FUNCTION_BLOCK Agua_Reuso_HMI (* Service Interface Function Block Type *)
  (* Standard: 61499-2 *)
  (* Version 1.2, 15/10/2026, Hidryco, Hidryco, IHM da Agua_Reuso *)
  PACKAGE Hidryco.HidrycoLib;
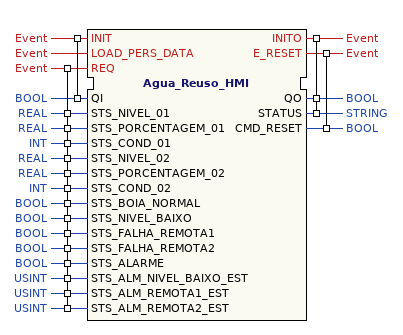
  EVENT_INPUT
    INIT WITH QI;
    LOAD_PERS_DATA; (* Reenvia os parametros persistentes *)
    REQ WITH STS_NIVEL_01, STS_PORCENTAGEM_01, STS_COND_01, STS_NIVEL_02, STS_PORCENTAGEM_02, STS_COND_02, STS_BOIA_NORMAL, STS_NIVEL_BAIXO, STS_FALHA_REMOTA1, STS_FALHA_REMOTA2, STS_ALARME, STS_ALM_NIVEL_BAIXO_EST, STS_ALM_REMOTA1_EST, STS_ALM_REMOTA2_EST; (* Atualizacao de status *)
  END_EVENT
  EVENT_OUTPUT
    INITO WITH QO, STATUS;
    E_RESET WITH CMD_RESET;
  END_EVENT
  VAR_INPUT
    QI : BOOL;
    STS_NIVEL_01 : REAL; (* Nivel 1000-PIT-01 *)
    STS_PORCENTAGEM_01 : REAL; (* Nivel 1000-PIT-01 (%) *)
    STS_COND_01 : INT; (* PIT-01: 0 normal, 1 HH, 2 H, 3 L, 4 LL, 5 sinal invalido, 6 falha memorizada, 7 desabilitado *)
    STS_NIVEL_02 : REAL; (* Nivel 1000-PIT-02 *)
    STS_PORCENTAGEM_02 : REAL; (* Nivel 1000-PIT-02 (%) *)
    STS_COND_02 : INT; (* PIT-02: mesmos codigos do STS_COND_01 *)
    STS_BOIA_NORMAL : BOOL; (* Boia 1000-LSL-01 levantada *)
    STS_NIVEL_BAIXO : BOOL; (* Nivel baixo pela boia 1000-LSL-01 *)
    STS_FALHA_REMOTA1 : BOOL; (* Falha de comunicacao com a remota 1 da Subestacao *)
    STS_FALHA_REMOTA2 : BOOL; (* Falha de comunicacao com a remota 2 da Subestacao *)
    STS_ALARME : BOOL; (* Algum alarme da agua de reuso *)
    STS_ALM_NIVEL_BAIXO_EST : USINT; (* Estado do ALARM_BIT nivel baixo (boia) (0 normal, 1 ativo reconhecido, 2 ativo nao reconhecido, 3 saiu nao reconhecido, 4 ativo e saiu nao reconhecido) *)
    STS_ALM_REMOTA1_EST : USINT; (* Estado do ALARM_BIT remota 1 (0 normal, 1 ativo reconhecido, 2 ativo nao reconhecido, 3 saiu nao reconhecido, 4 ativo e saiu nao reconhecido) *)
    STS_ALM_REMOTA2_EST : USINT; (* Estado do ALARM_BIT remota 2 (0 normal, 1 ativo reconhecido, 2 ativo nao reconhecido, 3 saiu nao reconhecido, 4 ativo e saiu nao reconhecido) *)
  END_VAR
  VAR_OUTPUT
    QO : BOOL; (* Event Output Qualifier *)
    STATUS : STRING; (* Service Status *)
    CMD_RESET : BOOL; (* Reconhece os alarmes da agua de reuso e faz o reset dos sensores *)
  END_VAR
  SERVICE /
    SEQUENCE 
    END_SEQUENCE
  END_SERVICE
END_FUNCTION_BLOCK
